// TIA Portal V20 export
FUNCTION_BLOCK "03_Betriebsart"   // FB16, LAD
{ S7_Optimized_Access := 'TRUE' }
// stored: MemoryReserve 100, SetENOAutomatically false
   VAR
      Projektnummer : WString;   // Projektnummer
      Projektname : WString;   // Projektname
      Validierung_Datum : WString;   // Datum an dem die Validierung ausgeführt wurde
      Validierung_Name : WString;   // Name der Person die die Validierung durchgeführt hat
      Validierung_F_PROG_SIG : DWord;   // F-Gesamtsignatur des Sicherheitsprogramms am Tag der Validierung
      Aktuell_F_PROG_SIG : DWord;   // Aktuelle F-Gesamtsignatur des Sicherheitsprogramms
      F_PROG_SIG_stimmt_überein : Bool;   // Aktuelle F-Gesamtsignatur stimmt mit der F-Gesamtsignatur am Tag der Validierung überein
      Simulation_aktiv : Bool;   // Simulation Software aktiv
      IN_Betriebsart_Manuell { ExternalAccessible := 'False'; ExternalVisible := 'False'; ExternalWritable := 'False'} : Bool;
      BA_Automatik_HMFP : Bool;   // Betriebsart Automatik Hilfsvariable Flanke
      BA_Automatik_FP : Bool;   // Betriebsart Automatik Flanke positiv
      IN_Betriebsart_Automatik { ExternalAccessible := 'False'; ExternalVisible := 'False'; ExternalWritable := 'False'} : Bool;
      BA_Verwaltung_HMFP : Bool;   // Betriebsart Verwaltung Hilfsvariable Flanke
      BA_Verwaltung_FP : Bool;   // Betriebsart Verwaltung Flanke positiv
      IN_Betriebsart_Verwaltung { ExternalAccessible := 'False'; ExternalVisible := 'False'; ExternalWritable := 'False'} : Bool;
      IN_Betriebsart_Richten { ExternalAccessible := 'False'; ExternalVisible := 'False'; ExternalWritable := 'False'} : Bool;
      Systemdruck_OK : Bool;
      Betriebsart : Int;   // Betriebsart 0= AUS, 1 = Manuell, 2=Automatik, 3= Verwaltung, 4= Richten
      BA_Manuell_HMFP : Bool;   // Betriebsart Manuell Hilfsvariable Flanke
      BA_Manuell_FP : Bool;   // Betriebsart Manuell Flanke positiv
      BA_Manuell : Bool;
      BA_Automatik : Bool;
      BA_Verwaltung : Bool;
      BA_Richten_HMFP : Bool;   // Betriebsart Richten Hilfsvariable Flanke
      BA_Richten_FP : Bool;   // Betriebsart Richten Flanke positiv
      BA_Richten : Bool;
      BA_0 : Bool;
      BA_0_HMFP : Bool;   // Betriebsart 0 Hilfsvariable Flanke
      BA_0_FP : Bool;   // Betriebsart 0 Flanke positiv
      BA_0_groesser_1_5 : Bool;
      TON_BA_0_groesser_1_5 { S7_SetPoint := 'True'} : TON_TIME;
      TON_Rücksetzen_der_Betriebsart { S7_SetPoint := 'True'} : TON_TIME;
      TON_Türen_setzen_zum_öffnen { S7_SetPoint := 'True'} : TON_TIME;
      "TOF_MRW Not-Halt Überwachung deaktivieren" { S7_SetPoint := 'True'} : TOF_TIME;
      HM_MRW_Zeitverzögerung { S7_SetPoint := 'True'} : Bool;   // Schutztüren sind verriegelt
      Türen_sind_verriegelt { S7_SetPoint := 'True'} : Bool;
      "NOT-HALT OK" : Bool;
      "NOT-HALT_HMFN" : Bool;   // NOT-HALT Hilfsvariable Flanke
      "NOT-HALT_FN" : Bool;   // NOT-HALT Flanke Negativ -> NOT-HALT hat ausgelöst
      Start_Taste : Bool;
      Start_Taste_HMFP : Bool;   // Start-Taste Hilfsvariable Flanke
      Start_Taste_FP : Bool;   // Start-Taste Flanke positiv
      ACK_Taste : Bool;
      ACK_Taste_HMFP : Bool;   // Start-Taste Flanke positiv
      ACK_Taste_FP : Bool;
      Stopp_Taste : Bool;
      "Schutztüren OK" : Bool;
      Schutztüren_HMFN : Bool;   // Schutztüren verriegelt Hilfsvariable Flanke
      Schutztüren_FN : Bool;   // Schutztüren verriegelt Flanke negativ
      Schutztüren_HMFP : Bool;   // Schutztüren verriegelt Hilfsvariable Flanke positiv
      Schutztüren_FP : Bool;   // Schutztüren verriegelt Flanke positiv
      "Druckbereich entlüftet" : Bool;
      Antriebe_sicher : Bool;
      Zuhaltung_Freigeben : Bool;
      Roboter_Motor_Ein : Bool;
      "P_Trig_Betriebsart Manuell" : Bool;
      "P_Trig_Betriebsart Automatik" : Bool;
      "P_Trig_Betriebsart Verwaltung" : Bool;
      "P_Trig_Betriebsart Richten" : Bool;
      TON_Hauptventil_aus { S7_SetPoint := 'True'} : TON_TIME;
      TON_Hauptventil_aus_status_Reset { S7_SetPoint := 'True'} : TON_TIME;
      Flanke_Hauptventil_aus { S7_SetPoint := 'True'} : Bool;
      Hauptventil_Reset : Bool;
      KP8_Bedienerkonsole { S7_SetPoint := 'True'} : "KP8";
   END_VAR
   VAR_TEMP
      TEMP_SK_Aktiv : Bool;
   END_VAR
   VAR_TEMP   // added for the SCL form of the ladder/FBD networks
      _w1 : Bool;
      _w2 : Bool;
      _w3 : Bool;
   END_VAR
BEGIN

REGION Network 1 (SCL): Projektinformationen

   #Projektnummer := WSTRING#'Au0199';
   #Projektname := WSTRING#'Steckzyklen Rotation';

   #Validierung_Datum := WSTRING#'18.06.2026';
   #Validierung_Name := WSTRING#'###';
   #Validierung_F_PROG_SIG := DW#16#C7164B37;   // F-Gesamtsignatur des Sicherheitsprogramms bei der Validierung
   (* D8254E31 *)
   #Aktuell_F_PROG_SIG := "RTG1SysInfo".F_SYSINFO.F_PROG_SIG; // F-Gesamtsignatur aktuell

   // Aktuelle F-Gesamtsignatur stimmt mit der F-Gesamtsignatur am Tag der Validierung überein
   IF #Aktuell_F_PROG_SIG = #Validierung_F_PROG_SIG THEN
       #F_PROG_SIG_stimmt_überein := true;
   ELSE
       #F_PROG_SIG_stimmt_überein := false;
   END_IF;
END_REGION

REGION Network 2 (SCL): Simulation Software

   #Simulation_aktiv := FALSE;
END_REGION

NETWORK
TITLE = Steuersignale Betriebsarten zuweisen
      A     "DE_Bedienerkonsole_Taste_K6_Manuell";
      =     #IN_Betriebsart_Manuell;

      A     "DE_Bedienerkonsole Taste_K7_Automatik";
      =     #IN_Betriebsart_Automatik;


      A     "DE_Bedienerkonsole_Taste_K4_Verwaltung";
      =     #IN_Betriebsart_Verwaltung;

      A     "DE_Bedienerkonsole_Taste_K5_Richten";
      =     #IN_Betriebsart_Richten;


      A     #BA_Richten;
      A     "DE_Bedienerkonsole_Taste_K3_Start";
      S     "HMI_COM".Richten_Gesamtanlage;



REGION Network 4: Systemdruck OK
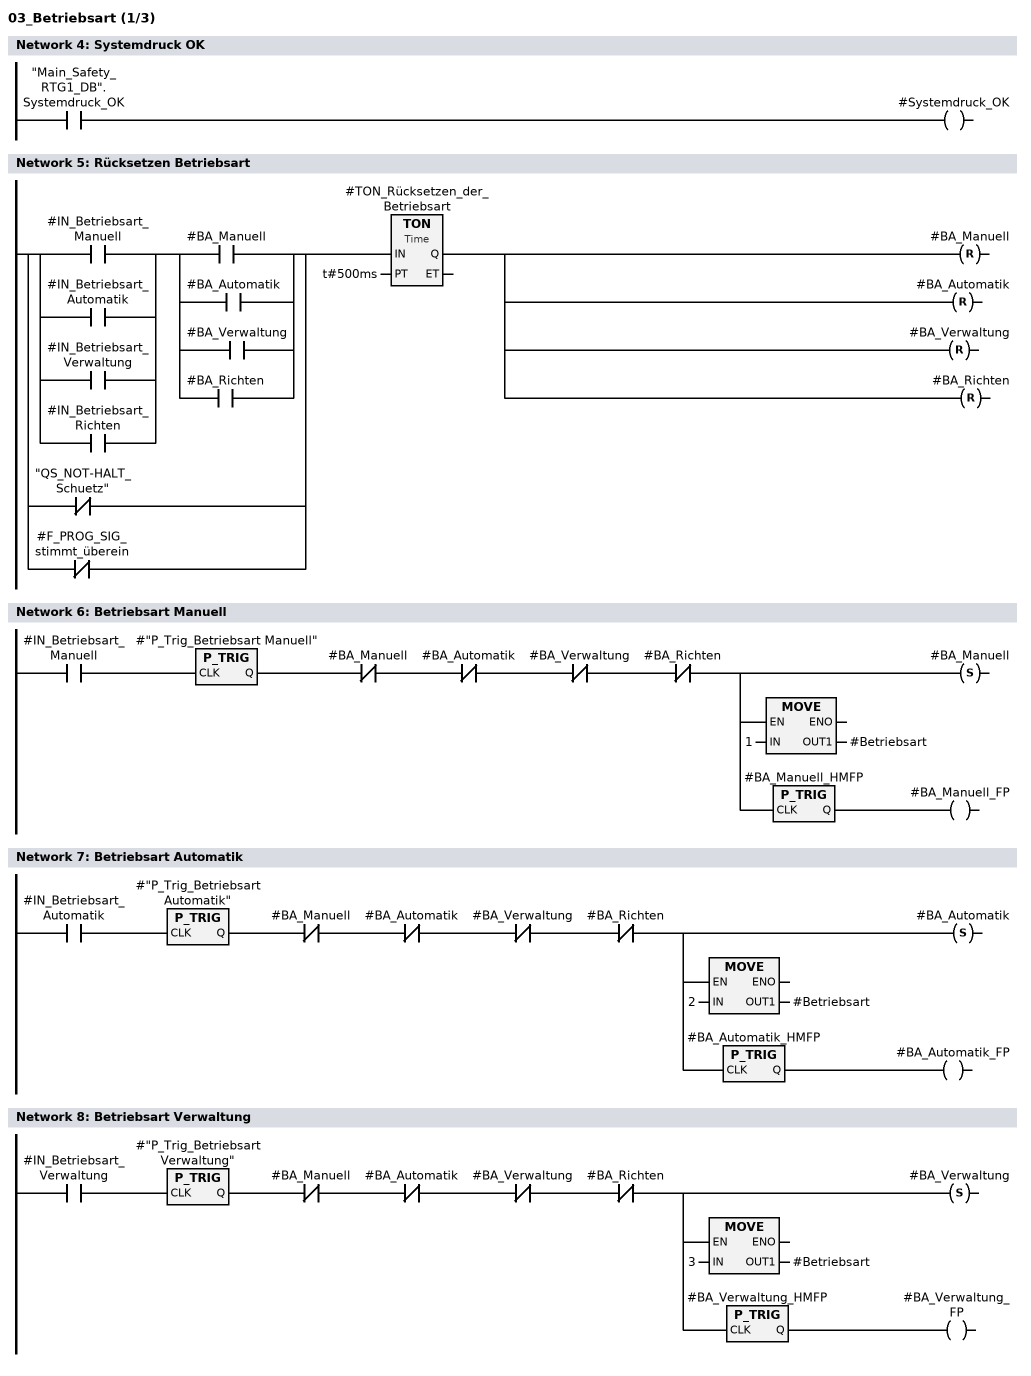
   RUNG wire#powerrail
      Contact( "Main_Safety_RTG1_DB".Systemdruck_OK )
      Coil( #Systemdruck_OK )
   END_RUNG
   // the same network as SCL:
   #Systemdruck_OK := "Main_Safety_RTG1_DB".Systemdruck_OK;
END_REGION

REGION Network 5: Rücksetzen Betriebsart
   RUNG wire#powerrail
      Contact( #IN_Betriebsart_Manuell )
      wire#w1
      Contact( #BA_Manuell )
      wire#w2
      { S7_Templates := "time_type := Time" } #TON_Rücksetzen_der_Betriebsart.TON(pt := t#500ms, et =>)
      wire#w3
      R_Coil( #BA_Manuell )
   END_RUNG
   RUNG wire#powerrail
      Contact( #IN_Betriebsart_Automatik )
   END_RUNG wire#w1
   RUNG wire#powerrail
      Contact( #IN_Betriebsart_Verwaltung )
   END_RUNG wire#w1
   RUNG wire#powerrail
      Contact( #IN_Betriebsart_Richten )
   END_RUNG wire#w1
   RUNG wire#w1
      Contact( #BA_Automatik )
   END_RUNG wire#w2
   RUNG wire#w1
      Contact( #BA_Verwaltung )
   END_RUNG wire#w2
   RUNG wire#w1
      Contact( #BA_Richten )
   END_RUNG wire#w2
   RUNG wire#powerrail
      I_Contact( "QS_NOT-HALT_Schuetz" )
   END_RUNG wire#w2
   RUNG wire#powerrail
      I_Contact( #F_PROG_SIG_stimmt_überein )
   END_RUNG wire#w2
   RUNG wire#w3
      R_Coil( #BA_Automatik )
   END_RUNG
   RUNG wire#w3
      R_Coil( #BA_Verwaltung )
   END_RUNG
   RUNG wire#w3
      R_Coil( #BA_Richten )
   END_RUNG
   // the same network as SCL:
   #TON_Rücksetzen_der_Betriebsart(IN := ((#IN_Betriebsart_Manuell OR #IN_Betriebsart_Automatik OR #IN_Betriebsart_Verwaltung OR #IN_Betriebsart_Richten) AND (#BA_Manuell OR #BA_Automatik OR #BA_Verwaltung OR #BA_Richten)) OR NOT "QS_NOT-HALT_Schuetz" OR NOT #F_PROG_SIG_stimmt_überein,   // TON
                           PT := t#500ms);
   IF #TON_Rücksetzen_der_Betriebsart.Q THEN
       #BA_Manuell := FALSE;
       #BA_Automatik := FALSE;
       #BA_Verwaltung := FALSE;
       #BA_Richten := FALSE;
   END_IF;
END_REGION

REGION Network 6: Betriebsart Manuell
   RUNG wire#powerrail
      Contact( #IN_Betriebsart_Manuell )
      P_Trig( #"P_Trig_Betriebsart Manuell" )
      I_Contact( #BA_Manuell )
      I_Contact( #BA_Automatik )
      I_Contact( #BA_Verwaltung )
      I_Contact( #BA_Richten )
      wire#w1
      S_Coil( #BA_Manuell )
   END_RUNG
   RUNG wire#w1
      Move(in := 1, out1 => #Betriebsart)
   END_RUNG
   RUNG wire#w1
      P_Trig( #BA_Manuell_HMFP )
      Coil( #BA_Manuell_FP )
   END_RUNG
   // the same network as SCL:
   #_w1 := #IN_Betriebsart_Manuell AND NOT #"P_Trig_Betriebsart Manuell";   // rising edge
   #"P_Trig_Betriebsart Manuell" := #IN_Betriebsart_Manuell;
   #_w2 := #_w1 AND NOT #BA_Manuell AND NOT #BA_Automatik AND NOT #BA_Verwaltung AND NOT #BA_Richten;
   IF #_w2 THEN
       #BA_Manuell := TRUE;
       #Betriebsart := 1;
   END_IF;
   #_w3 := #_w2 AND NOT #BA_Manuell_HMFP;   // rising edge
   #BA_Manuell_HMFP := #_w2;
   #BA_Manuell_FP := #_w3;
END_REGION

REGION Network 7: Betriebsart Automatik
   RUNG wire#powerrail
      Contact( #IN_Betriebsart_Automatik )
      P_Trig( #"P_Trig_Betriebsart Automatik" )
      I_Contact( #BA_Manuell )
      I_Contact( #BA_Automatik )
      I_Contact( #BA_Verwaltung )
      I_Contact( #BA_Richten )
      wire#w1
      S_Coil( #BA_Automatik )
   END_RUNG
   RUNG wire#w1
      Move(in := 2, out1 => #Betriebsart)
   END_RUNG
   RUNG wire#w1
      P_Trig( #BA_Automatik_HMFP )
      Coil( #BA_Automatik_FP )
   END_RUNG
   // the same network as SCL:
   #_w1 := #IN_Betriebsart_Automatik AND NOT #"P_Trig_Betriebsart Automatik";   // rising edge
   #"P_Trig_Betriebsart Automatik" := #IN_Betriebsart_Automatik;
   #_w2 := #_w1 AND NOT #BA_Manuell AND NOT #BA_Automatik AND NOT #BA_Verwaltung AND NOT #BA_Richten;
   IF #_w2 THEN
       #BA_Automatik := TRUE;
       #Betriebsart := 2;
   END_IF;
   #_w3 := #_w2 AND NOT #BA_Automatik_HMFP;   // rising edge
   #BA_Automatik_HMFP := #_w2;
   #BA_Automatik_FP := #_w3;
END_REGION

REGION Network 8: Betriebsart Verwaltung
   RUNG wire#powerrail
      Contact( #IN_Betriebsart_Verwaltung )
      P_Trig( #"P_Trig_Betriebsart Verwaltung" )
      I_Contact( #BA_Manuell )
      I_Contact( #BA_Automatik )
      I_Contact( #BA_Verwaltung )
      I_Contact( #BA_Richten )
      wire#w1
      S_Coil( #BA_Verwaltung )
   END_RUNG
   RUNG wire#w1
      Move(in := 3, out1 => #Betriebsart)
   END_RUNG
   RUNG wire#w1
      P_Trig( #BA_Verwaltung_HMFP )
      Coil( #BA_Verwaltung_FP )
   END_RUNG
   // the same network as SCL:
   #_w1 := #IN_Betriebsart_Verwaltung AND NOT #"P_Trig_Betriebsart Verwaltung";   // rising edge
   #"P_Trig_Betriebsart Verwaltung" := #IN_Betriebsart_Verwaltung;
   #_w2 := #_w1 AND NOT #BA_Manuell AND NOT #BA_Automatik AND NOT #BA_Verwaltung AND NOT #BA_Richten;
   IF #_w2 THEN
       #BA_Verwaltung := TRUE;
       #Betriebsart := 3;
   END_IF;
   #_w3 := #_w2 AND NOT #BA_Verwaltung_HMFP;   // rising edge
   #BA_Verwaltung_HMFP := #_w2;
   #BA_Verwaltung_FP := #_w3;
END_REGION

REGION Network 9: Betriebsart Richten
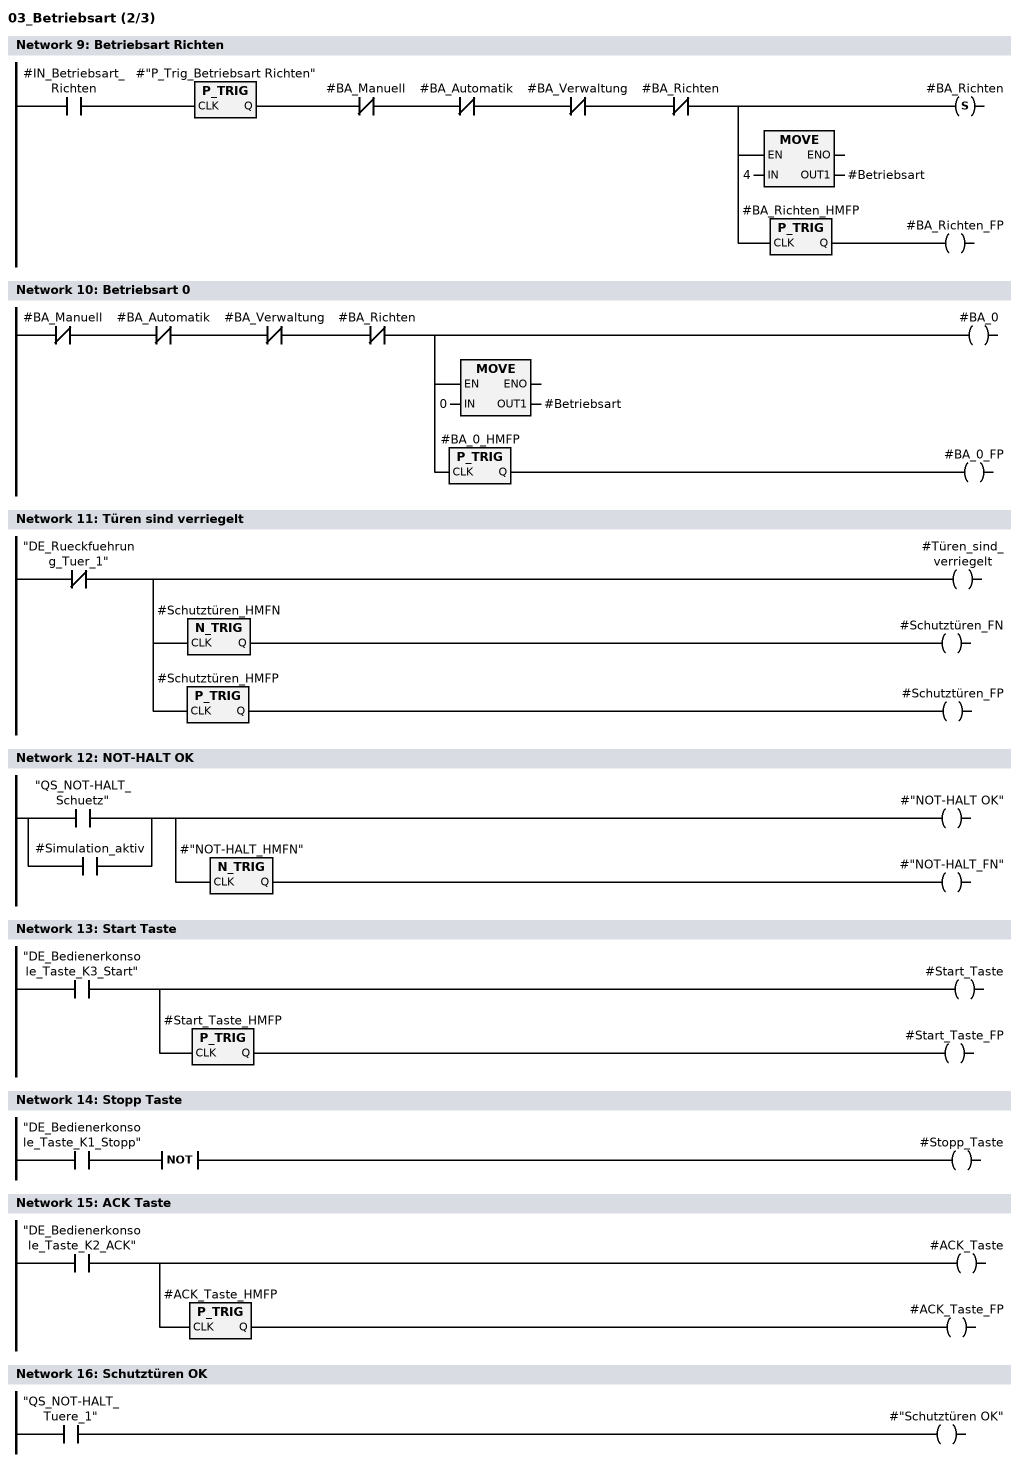
   RUNG wire#powerrail
      Contact( #IN_Betriebsart_Richten )
      P_Trig( #"P_Trig_Betriebsart Richten" )
      I_Contact( #BA_Manuell )
      I_Contact( #BA_Automatik )
      I_Contact( #BA_Verwaltung )
      I_Contact( #BA_Richten )
      wire#w1
      S_Coil( #BA_Richten )
   END_RUNG
   RUNG wire#w1
      Move(in := 4, out1 => #Betriebsart)
   END_RUNG
   RUNG wire#w1
      P_Trig( #BA_Richten_HMFP )
      Coil( #BA_Richten_FP )
   END_RUNG
   // the same network as SCL:
   #_w1 := #IN_Betriebsart_Richten AND NOT #"P_Trig_Betriebsart Richten";   // rising edge
   #"P_Trig_Betriebsart Richten" := #IN_Betriebsart_Richten;
   #_w2 := #_w1 AND NOT #BA_Manuell AND NOT #BA_Automatik AND NOT #BA_Verwaltung AND NOT #BA_Richten;
   IF #_w2 THEN
       #BA_Richten := TRUE;
       #Betriebsart := 4;
   END_IF;
   #_w3 := #_w2 AND NOT #BA_Richten_HMFP;   // rising edge
   #BA_Richten_HMFP := #_w2;
   #BA_Richten_FP := #_w3;
END_REGION

REGION Network 10: Betriebsart 0
   RUNG wire#powerrail
      I_Contact( #BA_Manuell )
      I_Contact( #BA_Automatik )
      I_Contact( #BA_Verwaltung )
      I_Contact( #BA_Richten )
      wire#w1
      Coil( #BA_0 )
   END_RUNG
   RUNG wire#w1
      Move(in := 0, out1 => #Betriebsart)
   END_RUNG
   RUNG wire#w1
      P_Trig( #BA_0_HMFP )
      Coil( #BA_0_FP )
   END_RUNG
   // the same network as SCL:
   #BA_0 := NOT #BA_Manuell AND NOT #BA_Automatik AND NOT #BA_Verwaltung AND NOT #BA_Richten;
   IF #BA_0 THEN #Betriebsart := 0; END_IF;
   #_w1 := #BA_0 AND NOT #BA_0_HMFP;   // rising edge
   #BA_0_HMFP := #BA_0;
   #BA_0_FP := #_w1;
END_REGION

REGION Network 11: Türen sind verriegelt
   RUNG wire#powerrail
      I_Contact( "DE_Rueckfuehrung_Tuer_1" )
      wire#w1
      Coil( #Türen_sind_verriegelt )
   END_RUNG
   RUNG wire#w1
      N_Trig( #Schutztüren_HMFN )
      Coil( #Schutztüren_FN )
   END_RUNG
   RUNG wire#w1
      P_Trig( #Schutztüren_HMFP )
      Coil( #Schutztüren_FP )
   END_RUNG
   // the same network as SCL:
   #Türen_sind_verriegelt := NOT "DE_Rueckfuehrung_Tuer_1";
   #_w1 := NOT (NOT "DE_Rueckfuehrung_Tuer_1") AND #Schutztüren_HMFN;   // falling edge
   #Schutztüren_HMFN := NOT "DE_Rueckfuehrung_Tuer_1";
   #Schutztüren_FN := #_w1;
   #_w2 := NOT "DE_Rueckfuehrung_Tuer_1" AND NOT #Schutztüren_HMFP;   // rising edge
   #Schutztüren_HMFP := NOT "DE_Rueckfuehrung_Tuer_1";
   #Schutztüren_FP := #_w2;
END_REGION

REGION Network 12: NOT-HALT OK
   RUNG wire#powerrail
      Contact( "QS_NOT-HALT_Schuetz" )
      wire#w1
      Coil( #"NOT-HALT OK" )
   END_RUNG
   RUNG wire#powerrail
      Contact( #Simulation_aktiv )
   END_RUNG wire#w1
   RUNG wire#w1
      N_Trig( #"NOT-HALT_HMFN" )
      Coil( #"NOT-HALT_FN" )
   END_RUNG
   // the same network as SCL:
   #"NOT-HALT OK" := "QS_NOT-HALT_Schuetz" OR #Simulation_aktiv;
   #_w1 := NOT #"NOT-HALT OK" AND #"NOT-HALT_HMFN";   // falling edge
   #"NOT-HALT_HMFN" := #"NOT-HALT OK";
   #"NOT-HALT_FN" := #_w1;
END_REGION

REGION Network 13: Start Taste
   RUNG wire#powerrail
      Contact( "DE_Bedienerkonsole_Taste_K3_Start" )
      wire#w1
      Coil( #Start_Taste )
   END_RUNG
   RUNG wire#w1
      P_Trig( #Start_Taste_HMFP )
      Coil( #Start_Taste_FP )
   END_RUNG
   // the same network as SCL:
   #Start_Taste := "DE_Bedienerkonsole_Taste_K3_Start";
   #_w1 := "DE_Bedienerkonsole_Taste_K3_Start" AND NOT #Start_Taste_HMFP;   // rising edge
   #Start_Taste_HMFP := "DE_Bedienerkonsole_Taste_K3_Start";
   #Start_Taste_FP := #_w1;
END_REGION

REGION Network 14: Stopp Taste
   RUNG wire#powerrail
      Contact( "DE_Bedienerkonsole_Taste_K1_Stopp" )
      Not()
      Coil( #Stopp_Taste )
   END_RUNG
   // the same network as SCL:
   #Stopp_Taste := NOT "DE_Bedienerkonsole_Taste_K1_Stopp";
END_REGION

REGION Network 15: ACK Taste
   RUNG wire#powerrail
      Contact( "DE_Bedienerkonsole_Taste_K2_ACK" )
      wire#w1
      Coil( #ACK_Taste )
   END_RUNG
   RUNG wire#w1
      P_Trig( #ACK_Taste_HMFP )
      Coil( #ACK_Taste_FP )
   END_RUNG
   // the same network as SCL:
   #ACK_Taste := "DE_Bedienerkonsole_Taste_K2_ACK";
   #_w1 := "DE_Bedienerkonsole_Taste_K2_ACK" AND NOT #ACK_Taste_HMFP;   // rising edge
   #ACK_Taste_HMFP := "DE_Bedienerkonsole_Taste_K2_ACK";
   #ACK_Taste_FP := #_w1;
END_REGION

REGION Network 16: Schutztüren OK
   RUNG wire#powerrail
      Contact( "QS_NOT-HALT_Tuere_1" )
      Coil( #"Schutztüren OK" )
   END_RUNG
   // the same network as SCL:
   #"Schutztüren OK" := "QS_NOT-HALT_Tuere_1";
END_REGION

REGION Network 17: Druckbereich entlüftet
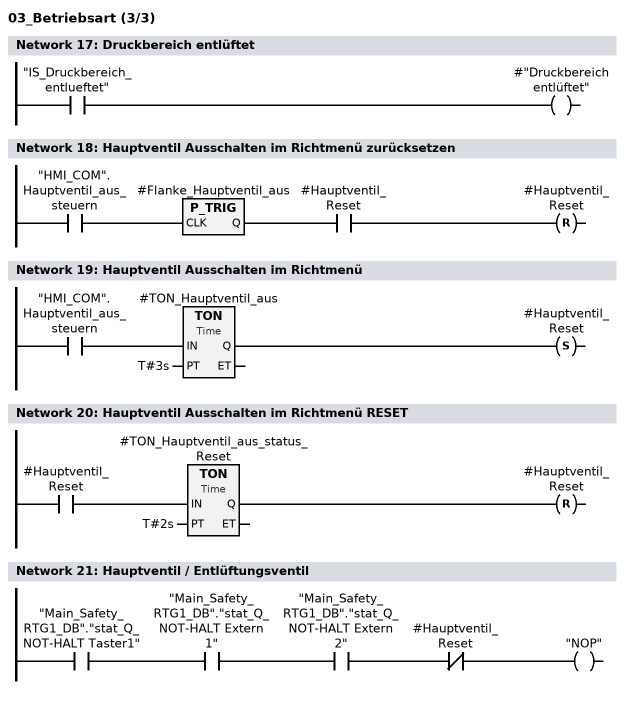
   RUNG wire#powerrail
      Contact( "IS_Druckbereich_entlueftet" )
      Coil( #"Druckbereich entlüftet" )
   END_RUNG
   // the same network as SCL:
   #"Druckbereich entlüftet" := "IS_Druckbereich_entlueftet";
END_REGION

REGION Network 18: Hauptventil Ausschalten im Richtmenü zurücksetzen
   RUNG wire#powerrail
      Contact( "HMI_COM".Hauptventil_aus_steuern )
      P_Trig( #Flanke_Hauptventil_aus )
      Contact( #Hauptventil_Reset )
      R_Coil( #Hauptventil_Reset )
   END_RUNG
   // the same network as SCL:
   #_w1 := "HMI_COM".Hauptventil_aus_steuern AND NOT #Flanke_Hauptventil_aus;   // rising edge
   #Flanke_Hauptventil_aus := "HMI_COM".Hauptventil_aus_steuern;
   IF #_w1 AND #Hauptventil_Reset THEN #Hauptventil_Reset := FALSE; END_IF;
END_REGION

REGION Network 19: Hauptventil Ausschalten im Richtmenü
   RUNG wire#powerrail
      Contact( "HMI_COM".Hauptventil_aus_steuern )
      { S7_Templates := "time_type := Time" } #TON_Hauptventil_aus.TON(pt := T#3s, et =>)
      S_Coil( #Hauptventil_Reset )
   END_RUNG
   // the same network as SCL:
   #TON_Hauptventil_aus(IN := "HMI_COM".Hauptventil_aus_steuern, PT := T#3s);   // TON
   IF #TON_Hauptventil_aus.Q THEN #Hauptventil_Reset := TRUE; END_IF;
END_REGION

REGION Network 20: Hauptventil Ausschalten im Richtmenü RESET
   RUNG wire#powerrail
      Contact( #Hauptventil_Reset )
      { S7_Templates := "time_type := Time" } #TON_Hauptventil_aus_status_Reset.TON(pt := T#2s, et =>)
      R_Coil( #Hauptventil_Reset )
   END_RUNG
   // the same network as SCL:
   #TON_Hauptventil_aus_status_Reset(IN := #Hauptventil_Reset, PT := T#2s);   // TON
   IF #TON_Hauptventil_aus_status_Reset.Q THEN #Hauptventil_Reset := FALSE; END_IF;
END_REGION

REGION Network 21: Hauptventil / Entlüftungsventil
   RUNG wire#powerrail
      Contact( "Main_Safety_RTG1_DB"."stat_Q_NOT-HALT Taster1" )
      Contact( "Main_Safety_RTG1_DB"."stat_Q_NOT-HALT Extern 1" )
      Contact( "Main_Safety_RTG1_DB"."stat_Q_NOT-HALT Extern 2" )
      I_Contact( #Hauptventil_Reset )
      Coil( "NOP" )
   END_RUNG
   // the same network as SCL:
   "NOP" := "Main_Safety_RTG1_DB"."stat_Q_NOT-HALT Taster1" AND "Main_Safety_RTG1_DB"."stat_Q_NOT-HALT Extern 1" AND "Main_Safety_RTG1_DB"."stat_Q_NOT-HALT Extern 2" AND NOT #Hauptventil_Reset;
END_REGION

NETWORK
TITLE = Flanke Takt 1.0
      A     "Clock_1Hz";
      FP    "HM_Clock_1Hz";
      =     "FL_Clock_1Hz";

NETWORK
TITLE = Status Signale LED
      A     "POS3_0_Signal".Station.SK_Aktiv;
      =     #TEMP_SK_Aktiv;

      CALL  #KP8_Bedienerkonsole
      ( IN_CLOCK           := "Clock_1Hz",
        IN_SAMMELSTÖRUNG   := "HMI_Signale".Sammelstoerung,
        IN_Grundstellung   := "HMI_COM".Grundstellung_Gesamt,
        IN_Ablauf_aktiv    := "HMI_Signale".Ablauf_aktiv,
        IN_Freigabe_Zyklus := "HMI_Signale".Freigabe_Zyklus,
        IN_SK_Aktiv        := #TEMP_SK_Aktiv,
        IN_BA_0            := #BA_0,
        IN_BA_RICHTEN      := #BA_Richten,
        IN_BA_MANUELL      := #BA_Manuell,
        IN_BA_AUTOMATIK    := #BA_Automatik,
        IN_BA_VERWALTUNG   := #BA_Verwaltung,
        AB_ROT             := "DA_Bedienerkonsole_Front_LED_K0-K7_ROT",
        AB_GRÜN            := "DA_Bedienerkonsole_Front_LED_K0-K7_GRÜN",
        AB_BLAU            := "DA_Bedienerkonsole_Front_LED_K0-K7_BLAU"
      );





END_FUNCTION_BLOCK
